(* IEC 61131-3 sources: trust-platform/examples/control/07-classical-stability-and-frequency-design/48-sensitivity-functions/src, 2 files *)

(* ---- Main.st ---- *)
USING Control;

(* Five periods of amplitude·sin(ω·t) from Start, then 0. *)
FUNCTION_BLOCK FivePeriodSine
VAR_INPUT
    Start : BOOL;
    Enable : BOOL;
    Amplitude : LREAL;
    OmegaRadS : LREAL;
END_VAR
VAR_OUTPUT
    Value : LREAL := 0.0;
    ElapsedS : LREAL := 0.0;
    Running : BOOL := FALSE;
END_VAR
IF Start THEN
    Running := TRUE;
    ElapsedS := LREAL#0.0;
END_IF;
IF NOT Enable THEN
    Running := FALSE;
END_IF;
IF Running AND ElapsedS >= LREAL#5.0 * LREAL#2.0 * LREAL#3.14159265358979 / OmegaRadS - LREAL#1.0E-9 THEN
    Running := FALSE;
END_IF;
IF Running THEN
    Value := Amplitude * SIN(OmegaRadS * ElapsedS);
    ElapsedS := ElapsedS + LREAL#0.1;
ELSE
    Value := LREAL#0.0;
END_IF;
END_FUNCTION_BLOCK

(* The loop transfer of this lesson, L = C·G with C = 5 + 1/s and G = 0.2·e^(−s)/(5s + 1): the PI zero cancels the
   heater's lag and L(jω) = 0.2·e^(−jω)/(jω) = −0.2·sin(ω)/ω − j·0.2·cos(ω)/ω. *)
FUNCTION LoopReal : LREAL
VAR_INPUT
    OmegaRadS : LREAL;
END_VAR
LoopReal := LREAL#-0.2 * SIN(OmegaRadS) / OmegaRadS;
END_FUNCTION

FUNCTION LoopImag : LREAL
VAR_INPUT
    OmegaRadS : LREAL;
END_VAR
LoopImag := LREAL#-0.2 * COS(OmegaRadS) / OmegaRadS;
END_FUNCTION

(* S = 1/(1 + L) and T = L/(1 + L). With 1 + L = a + jb, |S| = 1/√(a² + b²) and |T| = |L|·|S|. *)
FUNCTION SensitivityMagnitude : LREAL
VAR_INPUT
    LoopRealPart : LREAL;
    LoopImagPart : LREAL;
END_VAR
SensitivityMagnitude := LREAL#1.0 / SQRT((LREAL#1.0 + LoopRealPart) ** LREAL#2.0 + LoopImagPart ** LREAL#2.0);
END_FUNCTION

FUNCTION ComplementaryMagnitude : LREAL
VAR_INPUT
    LoopRealPart : LREAL;
    LoopImagPart : LREAL;
END_VAR
ComplementaryMagnitude := SQRT(LoopRealPart ** LREAL#2.0 + LoopImagPart ** LREAL#2.0)
    * SensitivityMagnitude(LoopRealPart := LoopRealPart, LoopImagPart := LoopImagPart);
END_FUNCTION

PROGRAM Main
VAR
    (* Two copies of the heater, each held at 35 °C by Control.PID as PI, Kp = 5 % per °C and Ki = 1 % per °C·s. *)
    LoadLoop : Control.PID;
    NoiseLoop : Control.PID;
    Parameters : Control.PIDParameters := (
        ProportionalGain := LREAL#5.0,
        IntegralGain := LREAL#1.0,
        DerivativeGain := LREAL#0.0,
        ProportionalSetpointWeight := LREAL#1.0,
        DerivativeSetpointWeight := LREAL#0.0,
        Bias := LREAL#0.0,
        OutputMinimum := LREAL#0.0,
        OutputMaximum := LREAL#100.0,
        RateMinimum := LREAL#-1000.0,
        RateMaximum := LREAL#1000.0,
        TrackingTime := LREAL#1.0,
        AntiWindup := PIDAntiWindup#BackCalculation
    );
    State : Control.PIDInitialState;
    LoadInput : Control.PIDInput;
    NoiseInput : Control.PIDInput;
    Initialized : BOOL := FALSE;
    SetpointC : LREAL := 35.0;
    (* The first heater: a heat load D enters the water. *)
    LoadTemperatureC : LREAL := 35.0;
    LoadCommandPct : LREAL := 75.0;
    LoadKw : LREAL := 0.0;
    (* The second heater: noise n enters only the reading its controller uses. *)
    NoiseTemperatureC : LREAL := 35.0;
    NoiseCommandPct : LREAL := 75.0;
    NoiseHeaterLoadKw : LREAL := 0.0;
    NoiseC : LREAL := 0.0;
    MeasuredTemperatureC : LREAL := 35.0;
    (* Control Studio's project experiment starts both injections: five periods at 0.2 rad/s. *)
    LoadSource : FivePeriodSine;
    NoiseSource : FivePeriodSine;
    LoadAmplitudeKw : LREAL := 10.0;
    NoiseAmplitudeC : LREAL := 0.05;
    OmegaRadS : LREAL := 0.2;
    ExperimentEnabled : BOOL := FALSE;
    ExperimentWasEnabled : BOOL := FALSE;
    Start : BOOL := FALSE;
    (* |S| and |T| at OmegaRadS. *)
    SensitivityAtOmega : LREAL := 0.0;
    ComplementaryAtOmega : LREAL := 0.0;
END_VAR

SensitivityAtOmega := SensitivityMagnitude(LoopRealPart := LoopReal(OmegaRadS := OmegaRadS),
    LoopImagPart := LoopImag(OmegaRadS := OmegaRadS));
ComplementaryAtOmega := ComplementaryMagnitude(LoopRealPart := LoopReal(OmegaRadS := OmegaRadS),
    LoopImagPart := LoopImag(OmegaRadS := OmegaRadS));

SetpointC := LREAL#35.0;
Start := ExperimentEnabled AND NOT ExperimentWasEnabled;
ExperimentWasEnabled := ExperimentEnabled;
LoadSource(Start := Start, Enable := ExperimentEnabled, Amplitude := LoadAmplitudeKw, OmegaRadS := OmegaRadS);
NoiseSource(Start := Start, Enable := ExperimentEnabled, Amplitude := NoiseAmplitudeC, OmegaRadS := OmegaRadS);
LoadKw := LoadSource.Value;
NoiseC := NoiseSource.Value;
NoiseHeaterLoadKw := LREAL#0.0;
MeasuredTemperatureC := NoiseTemperatureC + NoiseC;

LoadLoop.Configure(Parameters := Parameters);
NoiseLoop.Configure(Parameters := Parameters);
IF NOT Initialized THEN
    State.Setpoint := SetpointC;
    State.ProcessValue := SetpointC;
    State.NominalOutput := LREAL#75.0;
    State.SaturatedOutput := LREAL#75.0;
    LoadLoop.Initialize(State := State);
    NoiseLoop.Initialize(State := State);
    Initialized := TRUE;
END_IF;
LoadInput.Mode := PIDMode#Auto;
LoadInput.CycleTime := LREAL#0.1;
LoadInput.Setpoint := SetpointC;
LoadInput.ProcessValue := LoadTemperatureC;
LoadCommandPct := LoadLoop.Update(Input := LoadInput);
NoiseInput.Mode := PIDMode#Auto;
NoiseInput.CycleTime := LREAL#0.1;
NoiseInput.Setpoint := SetpointC;
NoiseInput.ProcessValue := MeasuredTemperatureC;
NoiseCommandPct := NoiseLoop.Update(Input := NoiseInput);
END_PROGRAM

CONFIGURATION Config
RESOURCE Res ON PLC
    TASK MainTask(INTERVAL := T#100ms, PRIORITY := 1);
    PROGRAM P1 WITH MainTask : Main;
END_RESOURCE
VAR_CONFIG
    P1.LoadCommandPct AT %QL0 : LREAL;
    P1.LoadKw AT %QL8 : LREAL;
    P1.NoiseCommandPct AT %QL16 : LREAL;
    P1.NoiseHeaterLoadKw AT %QL24 : LREAL;
    P1.LoadTemperatureC AT %IL0 : LREAL;
    P1.NoiseTemperatureC AT %IL8 : LREAL;
    P1.NoiseC AT %ML0 : LREAL;
    P1.MeasuredTemperatureC AT %ML8 : LREAL;
    P1.ExperimentEnabled AT %MX24.0 : BOOL;
    P1.SetpointC AT %ML16 : LREAL;
    P1.SensitivityAtOmega AT %ML32 : LREAL;
    P1.ComplementaryAtOmega AT %ML40 : LREAL;
END_VAR
END_CONFIGURATION

(* ---- tests.st ---- *)
(* @trustlsp:runtime-ignore — run these assertions with trust-dev test;
   they are not scheduled PLC instances in the lesson simulator. *)

TEST_PROGRAM TheLoopAtTheTestRate
(* L(j0.2) = −j·e^(−j0.2) = −sin 0.2 − j·cos 0.2: |L| = 1 at −101.46°. *)
ASSERT_NEAR(EXPECTED := LREAL#-0.198669, ACTUAL := LoopReal(OmegaRadS := LREAL#0.2), DELTA := LREAL#1.0e-6);
ASSERT_NEAR(EXPECTED := LREAL#-0.980067, ACTUAL := LoopImag(OmegaRadS := LREAL#0.2), DELTA := LREAL#1.0e-6);
END_TEST_PROGRAM

TEST_PROGRAM SensitivityAndComplement
VAR
    A : LREAL;
    B : LREAL;
    SReal : LREAL;
    SImag : LREAL;
    TReal : LREAL;
    TImag : LREAL;
END_VAR
(* |1 + L| = √(2 − 2·sin 0.2) = 1.26596, so |S| = |T| = 0.78991. *)
ASSERT_NEAR(EXPECTED := LREAL#0.78991, ACTUAL := SensitivityMagnitude(LoopRealPart := LoopReal(OmegaRadS := LREAL#0.2),
    LoopImagPart := LoopImag(OmegaRadS := LREAL#0.2)), DELTA := LREAL#1.0e-5);
ASSERT_NEAR(EXPECTED := LREAL#0.78991, ACTUAL := ComplementaryMagnitude(LoopRealPart := LoopReal(OmegaRadS := LREAL#0.2),
    LoopImagPart := LoopImag(OmegaRadS := LREAL#0.2)), DELTA := LREAL#1.0e-5);
(* S + T = 1 as complex numbers, yet |S| + |T| = 1.58. *)
A := LREAL#1.0 + LoopReal(OmegaRadS := LREAL#0.2);
B := LoopImag(OmegaRadS := LREAL#0.2);
SReal := A / (A * A + B * B);
SImag := -B / (A * A + B * B);
(* T = L/(1 + L) = L·(A − jB)/(A² + B²). *)
TReal := (LoopReal(OmegaRadS := LREAL#0.2) * A + LoopImag(OmegaRadS := LREAL#0.2) * B) / (A * A + B * B);
TImag := (LoopImag(OmegaRadS := LREAL#0.2) * A - LoopReal(OmegaRadS := LREAL#0.2) * B) / (A * A + B * B);
ASSERT_NEAR(EXPECTED := LREAL#1.0, ACTUAL := SReal + TReal, DELTA := LREAL#1.0e-12);
ASSERT_NEAR(EXPECTED := LREAL#0.0, ACTUAL := SImag + TImag, DELTA := LREAL#1.0e-12);
ASSERT_NEAR(EXPECTED := LREAL#1.57982, ACTUAL := SQRT(SReal * SReal + SImag * SImag) + SQRT(TReal * TReal + TImag * TImag), DELTA := LREAL#1.0e-5);
ASSERT_NEAR(EXPECTED := SQRT(SReal * SReal + SImag * SImag), ACTUAL := SensitivityMagnitude(LoopRealPart := LoopReal(OmegaRadS := LREAL#0.2),
    LoopImagPart := LoopImag(OmegaRadS := LREAL#0.2)), DELTA := LREAL#1.0e-12);
END_TEST_PROGRAM

TEST_PROGRAM ThePredictedAmplitudes
(* 10 kW load: 10·(0.1/√2)·|S| = 0.5586 °C. Noise 0.05 °C: water |T|·0.05 = 0.0395 °C, command |C|·|S|·0.05 = 0.2793 %. *)
ASSERT_NEAR(EXPECTED := LREAL#0.5586, ACTUAL := LREAL#10.0 * LREAL#0.1 / SQRT(LREAL#2.0)
    * SensitivityMagnitude(LoopRealPart := LoopReal(OmegaRadS := LREAL#0.2), LoopImagPart := LoopImag(OmegaRadS := LREAL#0.2)), DELTA := LREAL#1.0e-4);
ASSERT_NEAR(EXPECTED := LREAL#0.0395, ACTUAL := LREAL#0.05
    * ComplementaryMagnitude(LoopRealPart := LoopReal(OmegaRadS := LREAL#0.2), LoopImagPart := LoopImag(OmegaRadS := LREAL#0.2)), DELTA := LREAL#1.0e-4);
ASSERT_NEAR(EXPECTED := LREAL#0.2793, ACTUAL := LREAL#5.0 * SQRT(LREAL#2.0) * LREAL#0.05
    * SensitivityMagnitude(LoopRealPart := LoopReal(OmegaRadS := LREAL#0.2), LoopImagPart := LoopImag(OmegaRadS := LREAL#0.2)), DELTA := LREAL#1.0e-4);
END_TEST_PROGRAM
